DATA_BLOCK "GDB_LoadBankA"
{ S7_Optimized_Access := 'TRUE' }
VERSION : 0.1
NON_RETAIN
VAR
    Payload {ExternalAccessible := 'False'; ExternalVisible := 'False'; ExternalWritable := 'False'} : Array[0..63] of Byte;
END_VAR
BEGIN
END_DATA_BLOCK
